(* IEC 61131-3 sources: STAR-PLC-Agent/results/raw/codex_matrix_resume_20261114/codex_terra/SELF009/functional/attempt_0001, 1 file *)

(* ---- test_program.st ---- *)
PROGRAM PLC_PRG
VAR
 BenchStep : UDINT := 0;
 BenchCalls : UDINT := 0;
 BenchDone : BOOL := FALSE;
 BenchUut0 : FB_Task;
 BenchUut1 : FB_Task;
 BenchUut2 : FB_Task;
 BenchUut3 : FB_Task;
 BenchUut4 : FB_Task;
 BenchUut5 : FB_Task;
 BenchUut6 : FB_Task;
 TraceIn_PartPulse : ARRAY[0..55] OF BOOL;
 TraceIn_Reset : ARRAY[0..55] OF BOOL;
 TraceIn_Target : ARRAY[0..55] OF USINT;
 TraceOut_Count : ARRAY[0..55] OF USINT;
 TraceOut_Complete : ARRAY[0..55] OF BOOL;
 TraceOut_Error : ARRAY[0..55] OF BOOL;
END_VAR

IF NOT BenchDone THEN
 CASE BenchStep OF
 0:
   BenchUut0.PartPulse := FALSE;
   BenchUut0.Reset := FALSE;
   BenchUut0.Target := USINT#2;
   TraceIn_PartPulse[0] := BenchUut0.PartPulse;
   TraceIn_Reset[0] := BenchUut0.Reset;
   TraceIn_Target[0] := BenchUut0.Target;
   BenchUut0();
   TraceOut_Count[0] := BenchUut0.Count;
   TraceOut_Complete[0] := BenchUut0.Complete;
   TraceOut_Error[0] := BenchUut0.Error;
   BenchCalls := BenchCalls + 1;
 1:
   BenchUut0.PartPulse := TRUE;
   BenchUut0.Reset := FALSE;
   BenchUut0.Target := USINT#2;
   TraceIn_PartPulse[1] := BenchUut0.PartPulse;
   TraceIn_Reset[1] := BenchUut0.Reset;
   TraceIn_Target[1] := BenchUut0.Target;
   BenchUut0();
   TraceOut_Count[1] := BenchUut0.Count;
   TraceOut_Complete[1] := BenchUut0.Complete;
   TraceOut_Error[1] := BenchUut0.Error;
   BenchCalls := BenchCalls + 1;
 2:
   BenchUut0.PartPulse := TRUE;
   BenchUut0.Reset := FALSE;
   BenchUut0.Target := USINT#2;
   TraceIn_PartPulse[2] := BenchUut0.PartPulse;
   TraceIn_Reset[2] := BenchUut0.Reset;
   TraceIn_Target[2] := BenchUut0.Target;
   BenchUut0();
   TraceOut_Count[2] := BenchUut0.Count;
   TraceOut_Complete[2] := BenchUut0.Complete;
   TraceOut_Error[2] := BenchUut0.Error;
   BenchCalls := BenchCalls + 1;
 3:
   BenchUut0.PartPulse := FALSE;
   BenchUut0.Reset := FALSE;
   BenchUut0.Target := USINT#2;
   TraceIn_PartPulse[3] := BenchUut0.PartPulse;
   TraceIn_Reset[3] := BenchUut0.Reset;
   TraceIn_Target[3] := BenchUut0.Target;
   BenchUut0();
   TraceOut_Count[3] := BenchUut0.Count;
   TraceOut_Complete[3] := BenchUut0.Complete;
   TraceOut_Error[3] := BenchUut0.Error;
   BenchCalls := BenchCalls + 1;
 4:
   BenchUut0.PartPulse := TRUE;
   BenchUut0.Reset := FALSE;
   BenchUut0.Target := USINT#2;
   TraceIn_PartPulse[4] := BenchUut0.PartPulse;
   TraceIn_Reset[4] := BenchUut0.Reset;
   TraceIn_Target[4] := BenchUut0.Target;
   BenchUut0();
   TraceOut_Count[4] := BenchUut0.Count;
   TraceOut_Complete[4] := BenchUut0.Complete;
   TraceOut_Error[4] := BenchUut0.Error;
   BenchCalls := BenchCalls + 1;
 5:
   BenchUut0.PartPulse := FALSE;
   BenchUut0.Reset := FALSE;
   BenchUut0.Target := USINT#2;
   TraceIn_PartPulse[5] := BenchUut0.PartPulse;
   TraceIn_Reset[5] := BenchUut0.Reset;
   TraceIn_Target[5] := BenchUut0.Target;
   BenchUut0();
   TraceOut_Count[5] := BenchUut0.Count;
   TraceOut_Complete[5] := BenchUut0.Complete;
   TraceOut_Error[5] := BenchUut0.Error;
   BenchCalls := BenchCalls + 1;
 6:
   BenchUut0.PartPulse := TRUE;
   BenchUut0.Reset := FALSE;
   BenchUut0.Target := USINT#2;
   TraceIn_PartPulse[6] := BenchUut0.PartPulse;
   TraceIn_Reset[6] := BenchUut0.Reset;
   TraceIn_Target[6] := BenchUut0.Target;
   BenchUut0();
   TraceOut_Count[6] := BenchUut0.Count;
   TraceOut_Complete[6] := BenchUut0.Complete;
   TraceOut_Error[6] := BenchUut0.Error;
   BenchCalls := BenchCalls + 1;
 7:
   BenchUut1.PartPulse := TRUE;
   BenchUut1.Reset := TRUE;
   BenchUut1.Target := USINT#1;
   TraceIn_PartPulse[7] := BenchUut1.PartPulse;
   TraceIn_Reset[7] := BenchUut1.Reset;
   TraceIn_Target[7] := BenchUut1.Target;
   BenchUut1();
   TraceOut_Count[7] := BenchUut1.Count;
   TraceOut_Complete[7] := BenchUut1.Complete;
   TraceOut_Error[7] := BenchUut1.Error;
   BenchCalls := BenchCalls + 1;
 8:
   BenchUut1.PartPulse := TRUE;
   BenchUut1.Reset := FALSE;
   BenchUut1.Target := USINT#1;
   TraceIn_PartPulse[8] := BenchUut1.PartPulse;
   TraceIn_Reset[8] := BenchUut1.Reset;
   TraceIn_Target[8] := BenchUut1.Target;
   BenchUut1();
   TraceOut_Count[8] := BenchUut1.Count;
   TraceOut_Complete[8] := BenchUut1.Complete;
   TraceOut_Error[8] := BenchUut1.Error;
   BenchCalls := BenchCalls + 1;
 9:
   BenchUut1.PartPulse := FALSE;
   BenchUut1.Reset := FALSE;
   BenchUut1.Target := USINT#1;
   TraceIn_PartPulse[9] := BenchUut1.PartPulse;
   TraceIn_Reset[9] := BenchUut1.Reset;
   TraceIn_Target[9] := BenchUut1.Target;
   BenchUut1();
   TraceOut_Count[9] := BenchUut1.Count;
   TraceOut_Complete[9] := BenchUut1.Complete;
   TraceOut_Error[9] := BenchUut1.Error;
   BenchCalls := BenchCalls + 1;
 10:
   BenchUut1.PartPulse := TRUE;
   BenchUut1.Reset := FALSE;
   BenchUut1.Target := USINT#1;
   TraceIn_PartPulse[10] := BenchUut1.PartPulse;
   TraceIn_Reset[10] := BenchUut1.Reset;
   TraceIn_Target[10] := BenchUut1.Target;
   BenchUut1();
   TraceOut_Count[10] := BenchUut1.Count;
   TraceOut_Complete[10] := BenchUut1.Complete;
   TraceOut_Error[10] := BenchUut1.Error;
   BenchCalls := BenchCalls + 1;
 11:
   BenchUut1.PartPulse := TRUE;
   BenchUut1.Reset := FALSE;
   BenchUut1.Target := USINT#0;
   TraceIn_PartPulse[11] := BenchUut1.PartPulse;
   TraceIn_Reset[11] := BenchUut1.Reset;
   TraceIn_Target[11] := BenchUut1.Target;
   BenchUut1();
   TraceOut_Count[11] := BenchUut1.Count;
   TraceOut_Complete[11] := BenchUut1.Complete;
   TraceOut_Error[11] := BenchUut1.Error;
   BenchCalls := BenchCalls + 1;
 12:
   BenchUut1.PartPulse := TRUE;
   BenchUut1.Reset := FALSE;
   BenchUut1.Target := USINT#21;
   TraceIn_PartPulse[12] := BenchUut1.PartPulse;
   TraceIn_Reset[12] := BenchUut1.Reset;
   TraceIn_Target[12] := BenchUut1.Target;
   BenchUut1();
   TraceOut_Count[12] := BenchUut1.Count;
   TraceOut_Complete[12] := BenchUut1.Complete;
   TraceOut_Error[12] := BenchUut1.Error;
   BenchCalls := BenchCalls + 1;
 13:
   BenchUut2.PartPulse := TRUE;
   BenchUut2.Reset := FALSE;
   BenchUut2.Target := USINT#2;
   TraceIn_PartPulse[13] := BenchUut2.PartPulse;
   TraceIn_Reset[13] := BenchUut2.Reset;
   TraceIn_Target[13] := BenchUut2.Target;
   BenchUut2();
   TraceOut_Count[13] := BenchUut2.Count;
   TraceOut_Complete[13] := BenchUut2.Complete;
   TraceOut_Error[13] := BenchUut2.Error;
   BenchCalls := BenchCalls + 1;
 14:
   BenchUut2.PartPulse := FALSE;
   BenchUut2.Reset := FALSE;
   BenchUut2.Target := USINT#2;
   TraceIn_PartPulse[14] := BenchUut2.PartPulse;
   TraceIn_Reset[14] := BenchUut2.Reset;
   TraceIn_Target[14] := BenchUut2.Target;
   BenchUut2();
   TraceOut_Count[14] := BenchUut2.Count;
   TraceOut_Complete[14] := BenchUut2.Complete;
   TraceOut_Error[14] := BenchUut2.Error;
   BenchCalls := BenchCalls + 1;
 15:
   BenchUut2.PartPulse := TRUE;
   BenchUut2.Reset := FALSE;
   BenchUut2.Target := USINT#2;
   TraceIn_PartPulse[15] := BenchUut2.PartPulse;
   TraceIn_Reset[15] := BenchUut2.Reset;
   TraceIn_Target[15] := BenchUut2.Target;
   BenchUut2();
   TraceOut_Count[15] := BenchUut2.Count;
   TraceOut_Complete[15] := BenchUut2.Complete;
   TraceOut_Error[15] := BenchUut2.Error;
   BenchCalls := BenchCalls + 1;
 16:
   BenchUut2.PartPulse := FALSE;
   BenchUut2.Reset := FALSE;
   BenchUut2.Target := USINT#5;
   TraceIn_PartPulse[16] := BenchUut2.PartPulse;
   TraceIn_Reset[16] := BenchUut2.Reset;
   TraceIn_Target[16] := BenchUut2.Target;
   BenchUut2();
   TraceOut_Count[16] := BenchUut2.Count;
   TraceOut_Complete[16] := BenchUut2.Complete;
   TraceOut_Error[16] := BenchUut2.Error;
   BenchCalls := BenchCalls + 1;
 17:
   BenchUut2.PartPulse := FALSE;
   BenchUut2.Reset := FALSE;
   BenchUut2.Target := USINT#1;
   TraceIn_PartPulse[17] := BenchUut2.PartPulse;
   TraceIn_Reset[17] := BenchUut2.Reset;
   TraceIn_Target[17] := BenchUut2.Target;
   BenchUut2();
   TraceOut_Count[17] := BenchUut2.Count;
   TraceOut_Complete[17] := BenchUut2.Complete;
   TraceOut_Error[17] := BenchUut2.Error;
   BenchCalls := BenchCalls + 1;
 18:
   BenchUut2.PartPulse := TRUE;
   BenchUut2.Reset := FALSE;
   BenchUut2.Target := USINT#255;
   TraceIn_PartPulse[18] := BenchUut2.PartPulse;
   TraceIn_Reset[18] := BenchUut2.Reset;
   TraceIn_Target[18] := BenchUut2.Target;
   BenchUut2();
   TraceOut_Count[18] := BenchUut2.Count;
   TraceOut_Complete[18] := BenchUut2.Complete;
   TraceOut_Error[18] := BenchUut2.Error;
   BenchCalls := BenchCalls + 1;
 19:
   BenchUut2.PartPulse := TRUE;
   BenchUut2.Reset := FALSE;
   BenchUut2.Target := USINT#20;
   TraceIn_PartPulse[19] := BenchUut2.PartPulse;
   TraceIn_Reset[19] := BenchUut2.Reset;
   TraceIn_Target[19] := BenchUut2.Target;
   BenchUut2();
   TraceOut_Count[19] := BenchUut2.Count;
   TraceOut_Complete[19] := BenchUut2.Complete;
   TraceOut_Error[19] := BenchUut2.Error;
   BenchCalls := BenchCalls + 1;
 20:
   BenchUut2.PartPulse := FALSE;
   BenchUut2.Reset := FALSE;
   BenchUut2.Target := USINT#20;
   TraceIn_PartPulse[20] := BenchUut2.PartPulse;
   TraceIn_Reset[20] := BenchUut2.Reset;
   TraceIn_Target[20] := BenchUut2.Target;
   BenchUut2();
   TraceOut_Count[20] := BenchUut2.Count;
   TraceOut_Complete[20] := BenchUut2.Complete;
   TraceOut_Error[20] := BenchUut2.Error;
   BenchCalls := BenchCalls + 1;
 21:
   BenchUut2.PartPulse := TRUE;
   BenchUut2.Reset := FALSE;
   BenchUut2.Target := USINT#20;
   TraceIn_PartPulse[21] := BenchUut2.PartPulse;
   TraceIn_Reset[21] := BenchUut2.Reset;
   TraceIn_Target[21] := BenchUut2.Target;
   BenchUut2();
   TraceOut_Count[21] := BenchUut2.Count;
   TraceOut_Complete[21] := BenchUut2.Complete;
   TraceOut_Error[21] := BenchUut2.Error;
   BenchCalls := BenchCalls + 1;
 22:
   BenchUut3.PartPulse := FALSE;
   BenchUut3.Reset := FALSE;
   BenchUut3.Target := USINT#2;
   TraceIn_PartPulse[22] := BenchUut3.PartPulse;
   TraceIn_Reset[22] := BenchUut3.Reset;
   TraceIn_Target[22] := BenchUut3.Target;
   BenchUut3();
   TraceOut_Count[22] := BenchUut3.Count;
   TraceOut_Complete[22] := BenchUut3.Complete;
   TraceOut_Error[22] := BenchUut3.Error;
   BenchCalls := BenchCalls + 1;
 23:
   BenchUut3.PartPulse := TRUE;
   BenchUut3.Reset := FALSE;
   BenchUut3.Target := USINT#2;
   TraceIn_PartPulse[23] := BenchUut3.PartPulse;
   TraceIn_Reset[23] := BenchUut3.Reset;
   TraceIn_Target[23] := BenchUut3.Target;
   BenchUut3();
   TraceOut_Count[23] := BenchUut3.Count;
   TraceOut_Complete[23] := BenchUut3.Complete;
   TraceOut_Error[23] := BenchUut3.Error;
   BenchCalls := BenchCalls + 1;
 24:
   BenchUut3.PartPulse := TRUE;
   BenchUut3.Reset := FALSE;
   BenchUut3.Target := USINT#2;
   TraceIn_PartPulse[24] := BenchUut3.PartPulse;
   TraceIn_Reset[24] := BenchUut3.Reset;
   TraceIn_Target[24] := BenchUut3.Target;
   BenchUut3();
   TraceOut_Count[24] := BenchUut3.Count;
   TraceOut_Complete[24] := BenchUut3.Complete;
   TraceOut_Error[24] := BenchUut3.Error;
   BenchCalls := BenchCalls + 1;
 25:
   BenchUut3.PartPulse := FALSE;
   BenchUut3.Reset := FALSE;
   BenchUut3.Target := USINT#2;
   TraceIn_PartPulse[25] := BenchUut3.PartPulse;
   TraceIn_Reset[25] := BenchUut3.Reset;
   TraceIn_Target[25] := BenchUut3.Target;
   BenchUut3();
   TraceOut_Count[25] := BenchUut3.Count;
   TraceOut_Complete[25] := BenchUut3.Complete;
   TraceOut_Error[25] := BenchUut3.Error;
   BenchCalls := BenchCalls + 1;
 26:
   BenchUut3.PartPulse := TRUE;
   BenchUut3.Reset := FALSE;
   BenchUut3.Target := USINT#2;
   TraceIn_PartPulse[26] := BenchUut3.PartPulse;
   TraceIn_Reset[26] := BenchUut3.Reset;
   TraceIn_Target[26] := BenchUut3.Target;
   BenchUut3();
   TraceOut_Count[26] := BenchUut3.Count;
   TraceOut_Complete[26] := BenchUut3.Complete;
   TraceOut_Error[26] := BenchUut3.Error;
   BenchCalls := BenchCalls + 1;
 27:
   BenchUut3.PartPulse := FALSE;
   BenchUut3.Reset := FALSE;
   BenchUut3.Target := USINT#5;
   TraceIn_PartPulse[27] := BenchUut3.PartPulse;
   TraceIn_Reset[27] := BenchUut3.Reset;
   TraceIn_Target[27] := BenchUut3.Target;
   BenchUut3();
   TraceOut_Count[27] := BenchUut3.Count;
   TraceOut_Complete[27] := BenchUut3.Complete;
   TraceOut_Error[27] := BenchUut3.Error;
   BenchCalls := BenchCalls + 1;
 28:
   BenchUut4.PartPulse := TRUE;
   BenchUut4.Reset := FALSE;
   BenchUut4.Target := USINT#1;
   TraceIn_PartPulse[28] := BenchUut4.PartPulse;
   TraceIn_Reset[28] := BenchUut4.Reset;
   TraceIn_Target[28] := BenchUut4.Target;
   BenchUut4();
   TraceOut_Count[28] := BenchUut4.Count;
   TraceOut_Complete[28] := BenchUut4.Complete;
   TraceOut_Error[28] := BenchUut4.Error;
   BenchCalls := BenchCalls + 1;
 29:
   BenchUut4.PartPulse := TRUE;
   BenchUut4.Reset := FALSE;
   BenchUut4.Target := USINT#5;
   TraceIn_PartPulse[29] := BenchUut4.PartPulse;
   TraceIn_Reset[29] := BenchUut4.Reset;
   TraceIn_Target[29] := BenchUut4.Target;
   BenchUut4();
   TraceOut_Count[29] := BenchUut4.Count;
   TraceOut_Complete[29] := BenchUut4.Complete;
   TraceOut_Error[29] := BenchUut4.Error;
   BenchCalls := BenchCalls + 1;
 30:
   BenchUut4.PartPulse := FALSE;
   BenchUut4.Reset := FALSE;
   BenchUut4.Target := USINT#5;
   TraceIn_PartPulse[30] := BenchUut4.PartPulse;
   TraceIn_Reset[30] := BenchUut4.Reset;
   TraceIn_Target[30] := BenchUut4.Target;
   BenchUut4();
   TraceOut_Count[30] := BenchUut4.Count;
   TraceOut_Complete[30] := BenchUut4.Complete;
   TraceOut_Error[30] := BenchUut4.Error;
   BenchCalls := BenchCalls + 1;
 31:
   BenchUut4.PartPulse := TRUE;
   BenchUut4.Reset := FALSE;
   BenchUut4.Target := USINT#5;
   TraceIn_PartPulse[31] := BenchUut4.PartPulse;
   TraceIn_Reset[31] := BenchUut4.Reset;
   TraceIn_Target[31] := BenchUut4.Target;
   BenchUut4();
   TraceOut_Count[31] := BenchUut4.Count;
   TraceOut_Complete[31] := BenchUut4.Complete;
   TraceOut_Error[31] := BenchUut4.Error;
   BenchCalls := BenchCalls + 1;
 32:
   BenchUut4.PartPulse := TRUE;
   BenchUut4.Reset := FALSE;
   BenchUut4.Target := USINT#1;
   TraceIn_PartPulse[32] := BenchUut4.PartPulse;
   TraceIn_Reset[32] := BenchUut4.Reset;
   TraceIn_Target[32] := BenchUut4.Target;
   BenchUut4();
   TraceOut_Count[32] := BenchUut4.Count;
   TraceOut_Complete[32] := BenchUut4.Complete;
   TraceOut_Error[32] := BenchUut4.Error;
   BenchCalls := BenchCalls + 1;
 33:
   BenchUut4.PartPulse := TRUE;
   BenchUut4.Reset := FALSE;
   BenchUut4.Target := USINT#20;
   TraceIn_PartPulse[33] := BenchUut4.PartPulse;
   TraceIn_Reset[33] := BenchUut4.Reset;
   TraceIn_Target[33] := BenchUut4.Target;
   BenchUut4();
   TraceOut_Count[33] := BenchUut4.Count;
   TraceOut_Complete[33] := BenchUut4.Complete;
   TraceOut_Error[33] := BenchUut4.Error;
   BenchCalls := BenchCalls + 1;
 34:
   BenchUut4.PartPulse := TRUE;
   BenchUut4.Reset := FALSE;
   BenchUut4.Target := USINT#0;
   TraceIn_PartPulse[34] := BenchUut4.PartPulse;
   TraceIn_Reset[34] := BenchUut4.Reset;
   TraceIn_Target[34] := BenchUut4.Target;
   BenchUut4();
   TraceOut_Count[34] := BenchUut4.Count;
   TraceOut_Complete[34] := BenchUut4.Complete;
   TraceOut_Error[34] := BenchUut4.Error;
   BenchCalls := BenchCalls + 1;
 35:
   BenchUut4.PartPulse := TRUE;
   BenchUut4.Reset := FALSE;
   BenchUut4.Target := USINT#20;
   TraceIn_PartPulse[35] := BenchUut4.PartPulse;
   TraceIn_Reset[35] := BenchUut4.Reset;
   TraceIn_Target[35] := BenchUut4.Target;
   BenchUut4();
   TraceOut_Count[35] := BenchUut4.Count;
   TraceOut_Complete[35] := BenchUut4.Complete;
   TraceOut_Error[35] := BenchUut4.Error;
   BenchCalls := BenchCalls + 1;
 36:
   BenchUut4.PartPulse := FALSE;
   BenchUut4.Reset := FALSE;
   BenchUut4.Target := USINT#20;
   TraceIn_PartPulse[36] := BenchUut4.PartPulse;
   TraceIn_Reset[36] := BenchUut4.Reset;
   TraceIn_Target[36] := BenchUut4.Target;
   BenchUut4();
   TraceOut_Count[36] := BenchUut4.Count;
   TraceOut_Complete[36] := BenchUut4.Complete;
   TraceOut_Error[36] := BenchUut4.Error;
   BenchCalls := BenchCalls + 1;
 37:
   BenchUut4.PartPulse := TRUE;
   BenchUut4.Reset := FALSE;
   BenchUut4.Target := USINT#20;
   TraceIn_PartPulse[37] := BenchUut4.PartPulse;
   TraceIn_Reset[37] := BenchUut4.Reset;
   TraceIn_Target[37] := BenchUut4.Target;
   BenchUut4();
   TraceOut_Count[37] := BenchUut4.Count;
   TraceOut_Complete[37] := BenchUut4.Complete;
   TraceOut_Error[37] := BenchUut4.Error;
   BenchCalls := BenchCalls + 1;
 38:
   BenchUut5.PartPulse := FALSE;
   BenchUut5.Reset := FALSE;
   BenchUut5.Target := USINT#2;
   TraceIn_PartPulse[38] := BenchUut5.PartPulse;
   TraceIn_Reset[38] := BenchUut5.Reset;
   TraceIn_Target[38] := BenchUut5.Target;
   BenchUut5();
   TraceOut_Count[38] := BenchUut5.Count;
   TraceOut_Complete[38] := BenchUut5.Complete;
   TraceOut_Error[38] := BenchUut5.Error;
   BenchCalls := BenchCalls + 1;
 39:
   BenchUut5.PartPulse := TRUE;
   BenchUut5.Reset := FALSE;
   BenchUut5.Target := USINT#2;
   TraceIn_PartPulse[39] := BenchUut5.PartPulse;
   TraceIn_Reset[39] := BenchUut5.Reset;
   TraceIn_Target[39] := BenchUut5.Target;
   BenchUut5();
   TraceOut_Count[39] := BenchUut5.Count;
   TraceOut_Complete[39] := BenchUut5.Complete;
   TraceOut_Error[39] := BenchUut5.Error;
   BenchCalls := BenchCalls + 1;
 40:
   BenchUut5.PartPulse := TRUE;
   BenchUut5.Reset := FALSE;
   BenchUut5.Target := USINT#2;
   TraceIn_PartPulse[40] := BenchUut5.PartPulse;
   TraceIn_Reset[40] := BenchUut5.Reset;
   TraceIn_Target[40] := BenchUut5.Target;
   BenchUut5();
   TraceOut_Count[40] := BenchUut5.Count;
   TraceOut_Complete[40] := BenchUut5.Complete;
   TraceOut_Error[40] := BenchUut5.Error;
   BenchCalls := BenchCalls + 1;
 41:
   BenchUut5.PartPulse := FALSE;
   BenchUut5.Reset := FALSE;
   BenchUut5.Target := USINT#2;
   TraceIn_PartPulse[41] := BenchUut5.PartPulse;
   TraceIn_Reset[41] := BenchUut5.Reset;
   TraceIn_Target[41] := BenchUut5.Target;
   BenchUut5();
   TraceOut_Count[41] := BenchUut5.Count;
   TraceOut_Complete[41] := BenchUut5.Complete;
   TraceOut_Error[41] := BenchUut5.Error;
   BenchCalls := BenchCalls + 1;
 42:
   BenchUut5.PartPulse := TRUE;
   BenchUut5.Reset := FALSE;
   BenchUut5.Target := USINT#2;
   TraceIn_PartPulse[42] := BenchUut5.PartPulse;
   TraceIn_Reset[42] := BenchUut5.Reset;
   TraceIn_Target[42] := BenchUut5.Target;
   BenchUut5();
   TraceOut_Count[42] := BenchUut5.Count;
   TraceOut_Complete[42] := BenchUut5.Complete;
   TraceOut_Error[42] := BenchUut5.Error;
   BenchCalls := BenchCalls + 1;
 43:
   BenchUut5.PartPulse := FALSE;
   BenchUut5.Reset := FALSE;
   BenchUut5.Target := USINT#2;
   TraceIn_PartPulse[43] := BenchUut5.PartPulse;
   TraceIn_Reset[43] := BenchUut5.Reset;
   TraceIn_Target[43] := BenchUut5.Target;
   BenchUut5();
   TraceOut_Count[43] := BenchUut5.Count;
   TraceOut_Complete[43] := BenchUut5.Complete;
   TraceOut_Error[43] := BenchUut5.Error;
   BenchCalls := BenchCalls + 1;
 44:
   BenchUut5.PartPulse := TRUE;
   BenchUut5.Reset := FALSE;
   BenchUut5.Target := USINT#2;
   TraceIn_PartPulse[44] := BenchUut5.PartPulse;
   TraceIn_Reset[44] := BenchUut5.Reset;
   TraceIn_Target[44] := BenchUut5.Target;
   BenchUut5();
   TraceOut_Count[44] := BenchUut5.Count;
   TraceOut_Complete[44] := BenchUut5.Complete;
   TraceOut_Error[44] := BenchUut5.Error;
   BenchCalls := BenchCalls + 1;
 45:
   BenchUut5.PartPulse := FALSE;
   BenchUut5.Reset := FALSE;
   BenchUut5.Target := USINT#2;
   TraceIn_PartPulse[45] := BenchUut5.PartPulse;
   TraceIn_Reset[45] := BenchUut5.Reset;
   TraceIn_Target[45] := BenchUut5.Target;
   BenchUut5();
   TraceOut_Count[45] := BenchUut5.Count;
   TraceOut_Complete[45] := BenchUut5.Complete;
   TraceOut_Error[45] := BenchUut5.Error;
   BenchCalls := BenchCalls + 1;
 46:
   BenchUut5.PartPulse := FALSE;
   BenchUut5.Reset := FALSE;
   BenchUut5.Target := USINT#2;
   TraceIn_PartPulse[46] := BenchUut5.PartPulse;
   TraceIn_Reset[46] := BenchUut5.Reset;
   TraceIn_Target[46] := BenchUut5.Target;
   BenchUut5();
   TraceOut_Count[46] := BenchUut5.Count;
   TraceOut_Complete[46] := BenchUut5.Complete;
   TraceOut_Error[46] := BenchUut5.Error;
   BenchCalls := BenchCalls + 1;
 47:
   BenchUut6.PartPulse := FALSE;
   BenchUut6.Reset := FALSE;
   BenchUut6.Target := USINT#2;
   TraceIn_PartPulse[47] := BenchUut6.PartPulse;
   TraceIn_Reset[47] := BenchUut6.Reset;
   TraceIn_Target[47] := BenchUut6.Target;
   BenchUut6();
   TraceOut_Count[47] := BenchUut6.Count;
   TraceOut_Complete[47] := BenchUut6.Complete;
   TraceOut_Error[47] := BenchUut6.Error;
   BenchCalls := BenchCalls + 1;
 48:
   BenchUut6.PartPulse := TRUE;
   BenchUut6.Reset := FALSE;
   BenchUut6.Target := USINT#2;
   TraceIn_PartPulse[48] := BenchUut6.PartPulse;
   TraceIn_Reset[48] := BenchUut6.Reset;
   TraceIn_Target[48] := BenchUut6.Target;
   BenchUut6();
   TraceOut_Count[48] := BenchUut6.Count;
   TraceOut_Complete[48] := BenchUut6.Complete;
   TraceOut_Error[48] := BenchUut6.Error;
   BenchCalls := BenchCalls + 1;
 49:
   BenchUut6.PartPulse := TRUE;
   BenchUut6.Reset := FALSE;
   BenchUut6.Target := USINT#2;
   TraceIn_PartPulse[49] := BenchUut6.PartPulse;
   TraceIn_Reset[49] := BenchUut6.Reset;
   TraceIn_Target[49] := BenchUut6.Target;
   BenchUut6();
   TraceOut_Count[49] := BenchUut6.Count;
   TraceOut_Complete[49] := BenchUut6.Complete;
   TraceOut_Error[49] := BenchUut6.Error;
   BenchCalls := BenchCalls + 1;
 50:
   BenchUut6.PartPulse := FALSE;
   BenchUut6.Reset := FALSE;
   BenchUut6.Target := USINT#2;
   TraceIn_PartPulse[50] := BenchUut6.PartPulse;
   TraceIn_Reset[50] := BenchUut6.Reset;
   TraceIn_Target[50] := BenchUut6.Target;
   BenchUut6();
   TraceOut_Count[50] := BenchUut6.Count;
   TraceOut_Complete[50] := BenchUut6.Complete;
   TraceOut_Error[50] := BenchUut6.Error;
   BenchCalls := BenchCalls + 1;
 51:
   BenchUut6.PartPulse := TRUE;
   BenchUut6.Reset := FALSE;
   BenchUut6.Target := USINT#2;
   TraceIn_PartPulse[51] := BenchUut6.PartPulse;
   TraceIn_Reset[51] := BenchUut6.Reset;
   TraceIn_Target[51] := BenchUut6.Target;
   BenchUut6();
   TraceOut_Count[51] := BenchUut6.Count;
   TraceOut_Complete[51] := BenchUut6.Complete;
   TraceOut_Error[51] := BenchUut6.Error;
   BenchCalls := BenchCalls + 1;
 52:
   BenchUut6.PartPulse := FALSE;
   BenchUut6.Reset := FALSE;
   BenchUut6.Target := USINT#2;
   TraceIn_PartPulse[52] := BenchUut6.PartPulse;
   TraceIn_Reset[52] := BenchUut6.Reset;
   TraceIn_Target[52] := BenchUut6.Target;
   BenchUut6();
   TraceOut_Count[52] := BenchUut6.Count;
   TraceOut_Complete[52] := BenchUut6.Complete;
   TraceOut_Error[52] := BenchUut6.Error;
   BenchCalls := BenchCalls + 1;
 53:
   BenchUut6.PartPulse := TRUE;
   BenchUut6.Reset := FALSE;
   BenchUut6.Target := USINT#2;
   TraceIn_PartPulse[53] := BenchUut6.PartPulse;
   TraceIn_Reset[53] := BenchUut6.Reset;
   TraceIn_Target[53] := BenchUut6.Target;
   BenchUut6();
   TraceOut_Count[53] := BenchUut6.Count;
   TraceOut_Complete[53] := BenchUut6.Complete;
   TraceOut_Error[53] := BenchUut6.Error;
   BenchCalls := BenchCalls + 1;
 54:
   BenchUut6.PartPulse := TRUE;
   BenchUut6.Reset := TRUE;
   BenchUut6.Target := USINT#2;
   TraceIn_PartPulse[54] := BenchUut6.PartPulse;
   TraceIn_Reset[54] := BenchUut6.Reset;
   TraceIn_Target[54] := BenchUut6.Target;
   BenchUut6();
   TraceOut_Count[54] := BenchUut6.Count;
   TraceOut_Complete[54] := BenchUut6.Complete;
   TraceOut_Error[54] := BenchUut6.Error;
   BenchCalls := BenchCalls + 1;
 55:
   BenchUut6.PartPulse := TRUE;
   BenchUut6.Reset := TRUE;
   BenchUut6.Target := USINT#2;
   TraceIn_PartPulse[55] := BenchUut6.PartPulse;
   TraceIn_Reset[55] := BenchUut6.Reset;
   TraceIn_Target[55] := BenchUut6.Target;
   BenchUut6();
   TraceOut_Count[55] := BenchUut6.Count;
   TraceOut_Complete[55] := BenchUut6.Complete;
   TraceOut_Error[55] := BenchUut6.Error;
   BenchCalls := BenchCalls + 1;
 END_CASE;
 BenchStep := BenchStep + 1;
 IF BenchStep >= 56 THEN BenchDone := TRUE; END_IF;
END_IF;
END_PROGRAM
